(* IEC 61131-3 sources: rusty/tests/lit/single/exit, 39 files *)

(* ---- fb_exit_in_class.st ---- *)
// RUN: %COMPILE %s && %RUN | %CHECK %s
// A class can declare `FB_EXIT`. It runs for each instance when the application ends.
CLASS Logger
    METHOD FB_EXIT
        printf('logger$N');
    END_METHOD
END_CLASS

VAR_GLOBAL
    logger: Logger;
END_VAR

FUNCTION main: DINT
    printf('main done$N');
    // CHECK: main done
    // CHECK-NEXT: logger
    // CHECK-NOT: logger
END_FUNCTION

(* ---- array_elements_ascending.st ---- *)
// RUN: %COMPILE %s && %RUN | %CHECK %s
// The elements of an array are exited in ascending index order. The arrays themselves follow
// the reverse declaration order.
FUNCTION_BLOCK Slot
    VAR
        id: DINT;
    END_VAR

    METHOD FB_EXIT
        printf('slot %d$N', id);
    END_METHOD
END_FUNCTION_BLOCK

VAR_GLOBAL
    first: ARRAY[0..1] OF Slot := [(id := 1), (id := 2)];
    second: ARRAY[0..1] OF Slot := [(id := 3), (id := 4)];
END_VAR

FUNCTION main: DINT
    printf('main done$N');
    // CHECK: main done
    // CHECK-NEXT: slot 3
    // CHECK-NEXT: slot 4
    // CHECK-NEXT: slot 1
    // CHECK-NEXT: slot 2
    // CHECK-NOT: slot
END_FUNCTION

(* ---- array_with_negative_lower_bound.st ---- *)
// RUN: %COMPILE %s && %RUN | %CHECK %s
// An array whose range goes from a negative to a positive index is exited from its lowest
// index to its highest index. Each element prints its own index.
FUNCTION_BLOCK Slot
    VAR
        index: DINT;
    END_VAR

    METHOD FB_EXIT
        printf('slot %d$N', index);
    END_METHOD
END_FUNCTION_BLOCK

VAR_GLOBAL
    slots: ARRAY[-2..4] OF Slot;
END_VAR

FUNCTION main: DINT
    VAR
        i: DINT;
    END_VAR

    FOR i := -2 TO 4 DO
        slots[i].index := i;
    END_FOR

    printf('main done$N');
    // CHECK: main done
    // CHECK-NEXT: slot -2
    // CHECK-NEXT: slot -1
    // CHECK-NEXT: slot 0
    // CHECK-NEXT: slot 1
    // CHECK-NEXT: slot 2
    // CHECK-NEXT: slot 3
    // CHECK-NEXT: slot 4
    // CHECK-NOT: slot
END_FUNCTION

(* ---- array_with_two_dimensions.st ---- *)
// RUN: %COMPILE %s && %RUN | %CHECK %s
// The elements of an array with two dimensions are exited row by row: the last index changes
// first.
FUNCTION_BLOCK Slot
    VAR
        id: DINT;
    END_VAR

    METHOD FB_EXIT
        printf('slot %d$N', id);
    END_METHOD
END_FUNCTION_BLOCK

VAR_GLOBAL
    grid: ARRAY[1..2, 1..2] OF Slot;
END_VAR

FUNCTION main: DINT
    grid[1, 1].id := 11;
    grid[1, 2].id := 12;
    grid[2, 1].id := 21;
    grid[2, 2].id := 22;

    printf('main done$N');
    // CHECK: main done
    // CHECK-NEXT: slot 11
    // CHECK-NEXT: slot 12
    // CHECK-NEXT: slot 21
    // CHECK-NEXT: slot 22
    // CHECK-NOT: slot
END_FUNCTION

(* ---- container_before_members.st ---- *)
// RUN: %COMPILE %s && %RUN | %CHECK %s
// A function block runs its own `FB_EXIT` first, before any of its members is exited. The
// members follow in reverse declaration order.
FUNCTION_BLOCK Part
    VAR
        id: DINT;
    END_VAR

    METHOD FB_EXIT
        printf('part %d$N', id);
    END_METHOD
END_FUNCTION_BLOCK

FUNCTION_BLOCK Machine
    VAR
        first: Part := (id := 1);
        second: Part := (id := 2);
    END_VAR

    METHOD FB_EXIT
        printf('machine$N');
    END_METHOD
END_FUNCTION_BLOCK

VAR_GLOBAL
    machine: Machine;
END_VAR

FUNCTION main: DINT
    printf('main done$N');
    // CHECK: main done
    // CHECK-NEXT: machine
    // CHECK-NEXT: part 2
    // CHECK-NEXT: part 1
    // CHECK-NOT: {{machine|part}}
END_FUNCTION

(* ---- container_without_fb_exit.st ---- *)
// RUN: %COMPILE %s && %RUN | %CHECK %s
// A member is exited also when the function blocks that hold it declare no `FB_EXIT`, over
// more than one level.
FUNCTION_BLOCK Part
    METHOD FB_EXIT
        printf('part$N');
    END_METHOD
END_FUNCTION_BLOCK

FUNCTION_BLOCK Holder
    VAR
        part: Part;
    END_VAR
END_FUNCTION_BLOCK

FUNCTION_BLOCK Outer
    VAR
        holder: Holder;
    END_VAR
END_FUNCTION_BLOCK

VAR_GLOBAL
    outer: Outer;
END_VAR

FUNCTION main: DINT
    printf('main done$N');
    // CHECK: main done
    // CHECK-NEXT: part
    // CHECK-NOT: part
END_FUNCTION

(* ---- copy_by_assignment.st ---- *)
// RUN: %COMPILE %s && %RUN | %CHECK %s
// An assignment copies an instance with no call of `FB_INIT` or `FB_EXIT`. Each variable is
// exited one time, with the data it holds at that moment.
FUNCTION_BLOCK Token
    VAR
        id: DINT;
    END_VAR

    METHOD FB_EXIT
        printf('exit %d$N', id);
    END_METHOD
END_FUNCTION_BLOCK

VAR_GLOBAL
    target: Token := (id := 1);
    source: Token := (id := 2);
END_VAR

FUNCTION main: DINT
    target := source;
    printf('assigned$N');
    printf('main done$N');
    // CHECK: assigned
    // CHECK-NEXT: main done
    // CHECK-NEXT: exit 2
    // CHECK-NEXT: exit 2
    // CHECK-NOT: exit
END_FUNCTION

(* ---- copy_by_value_input.st ---- *)
// RUN: %COMPILE %s && %RUN | %CHECK %s
// An input that is passed by value is a copy of the argument, made with no call of `FB_INIT`.
// The copy is not exited at the end of the call. The argument is exited one time, when the
// application ends.
FUNCTION_BLOCK Token
    VAR
        id: DINT;
    END_VAR

    METHOD FB_EXIT
        printf('exit %d$N', id);
    END_METHOD
END_FUNCTION_BLOCK

FUNCTION inspect: DINT
    VAR_INPUT
        copy: Token;
    END_VAR

    printf('inspect %d$N', copy.id);
END_FUNCTION

VAR_GLOBAL
    source: Token := (id := 1);
END_VAR

FUNCTION main: DINT
    inspect(source);
    printf('main done$N');
    // CHECK: inspect 1
    // CHECK-NEXT: main done
    // CHECK-NEXT: exit 1
    // CHECK-NOT: exit
END_FUNCTION

(* ---- early_return_case.st ---- *)
// RUN: %COMPILE %s && %RUN | %CHECK %s
// A local instance is exited when the call leaves the body through a `RETURN` in a `CASE` branch.
// The statements after the `RETURN` do not run.
FUNCTION_BLOCK Guard
    METHOD FB_EXIT
        printf('exit$N');
    END_METHOD
END_FUNCTION_BLOCK

FUNCTION work: DINT
    VAR
        guard: Guard;
    END_VAR

    CASE 1 OF
        1: RETURN;
    END_CASE
    printf('not reached$N');
END_FUNCTION

FUNCTION main: DINT
    work();
    printf('main done$N');
    // CHECK-NOT: not reached
    // CHECK: exit
    // CHECK-NEXT: main done
    // CHECK-NOT: exit
END_FUNCTION

(* ---- early_return_for.st ---- *)
// RUN: %COMPILE %s && %RUN | %CHECK %s
// A local instance is exited when the call leaves the body through a `RETURN` in a `FOR` loop.
// The statements after the `RETURN` do not run.
FUNCTION_BLOCK Guard
    METHOD FB_EXIT
        printf('exit$N');
    END_METHOD
END_FUNCTION_BLOCK

FUNCTION work: DINT
    VAR
        guard: Guard;
        i: DINT;
    END_VAR

    FOR i := 0 TO 5 DO
        RETURN;
    END_FOR
    printf('not reached$N');
END_FUNCTION

FUNCTION main: DINT
    work();
    printf('main done$N');
    // CHECK-NOT: not reached
    // CHECK: exit
    // CHECK-NEXT: main done
    // CHECK-NOT: exit
END_FUNCTION

(* ---- early_return_if.st ---- *)
// RUN: %COMPILE %s && %RUN | %CHECK %s
// A local instance is exited when the call leaves the body through a `RETURN` in an `IF` branch.
// The statements after the `RETURN` do not run.
FUNCTION_BLOCK Guard
    METHOD FB_EXIT
        printf('exit$N');
    END_METHOD
END_FUNCTION_BLOCK

FUNCTION work: DINT
    VAR
        guard: Guard;
    END_VAR

    IF TRUE THEN
        RETURN;
    END_IF
    printf('not reached$N');
END_FUNCTION

FUNCTION main: DINT
    work();
    printf('main done$N');
    // CHECK-NOT: not reached
    // CHECK: exit
    // CHECK-NEXT: main done
    // CHECK-NOT: exit
END_FUNCTION

(* ---- early_return_repeat.st ---- *)
// RUN: %COMPILE %s && %RUN | %CHECK %s
// A local instance is exited when the call leaves the body through a `RETURN` in a `REPEAT` loop.
// The statements after the `RETURN` do not run.
FUNCTION_BLOCK Guard
    METHOD FB_EXIT
        printf('exit$N');
    END_METHOD
END_FUNCTION_BLOCK

FUNCTION work: DINT
    VAR
        guard: Guard;
    END_VAR

    REPEAT
        RETURN;
    UNTIL TRUE END_REPEAT
    printf('not reached$N');
END_FUNCTION

FUNCTION main: DINT
    work();
    printf('main done$N');
    // CHECK-NOT: not reached
    // CHECK: exit
    // CHECK-NEXT: main done
    // CHECK-NOT: exit
END_FUNCTION

(* ---- early_return_top_level.st ---- *)
// RUN: %COMPILE %s && %RUN | %CHECK %s
// A local instance is exited when the call leaves the body through a `RETURN` at the top level
// of the body. The statements after the `RETURN` do not run.
FUNCTION_BLOCK Guard
    METHOD FB_EXIT
        printf('exit$N');
    END_METHOD
END_FUNCTION_BLOCK

FUNCTION work: DINT
    VAR
        guard: Guard;
    END_VAR

    RETURN;
    printf('not reached$N');
END_FUNCTION

FUNCTION main: DINT
    work();
    printf('main done$N');
    // CHECK-NOT: not reached
    // CHECK: exit
    // CHECK-NEXT: main done
    // CHECK-NOT: exit
END_FUNCTION

(* ---- early_return_while.st ---- *)
// RUN: %COMPILE %s && %RUN | %CHECK %s
// A local instance is exited when the call leaves the body through a `RETURN` in a `WHILE` loop.
// The statements after the `RETURN` do not run.
FUNCTION_BLOCK Guard
    METHOD FB_EXIT
        printf('exit$N');
    END_METHOD
END_FUNCTION_BLOCK

FUNCTION work: DINT
    VAR
        guard: Guard;
    END_VAR

    WHILE TRUE DO
        RETURN;
    END_WHILE
    printf('not reached$N');
END_FUNCTION

FUNCTION main: DINT
    work();
    printf('main done$N');
    // CHECK-NOT: not reached
    // CHECK: exit
    // CHECK-NEXT: main done
    // CHECK-NOT: exit
END_FUNCTION

(* ---- explicit_call.st ---- *)
// RUN: %COMPILE %s && %RUN | %CHECK %s
// `FB_EXIT` is a normal method for user code. A call from user code runs it, and the call at
// the end of the application follows as usual.
FUNCTION_BLOCK Token
    VAR
        id: DINT;
    END_VAR

    METHOD FB_EXIT
        printf('exit %d$N', id);
    END_METHOD
END_FUNCTION_BLOCK

VAR_GLOBAL
    token: Token := (id := 1);
END_VAR

FUNCTION main: DINT
    token.FB_EXIT();
    printf('main done$N');
    // CHECK: exit 1
    // CHECK-NEXT: main done
    // CHECK-NEXT: exit 1
    // CHECK-NOT: exit
END_FUNCTION

(* ---- fb_exit_in_program.st ---- *)
// RUN: %COMPILE %s && %RUN | %CHECK %s
// A program can declare `FB_EXIT`. It runs when the application ends, before the members of the
// program are exited.
FUNCTION_BLOCK Part
    METHOD FB_EXIT
        printf('part$N');
    END_METHOD
END_FUNCTION_BLOCK

PROGRAM prog
    VAR
        part: Part;
    END_VAR

    METHOD FB_EXIT
        printf('prog$N');
    END_METHOD
END_PROGRAM

FUNCTION main: DINT
    printf('main done$N');
    // CHECK: main done
    // CHECK-NEXT: prog
    // CHECK-NEXT: part
    // CHECK-NOT: {{prog|part}}
END_FUNCTION

(* ---- function_locals.st ---- *)
// RUN: %COMPILE %s && %RUN | %CHECK %s
// A function block instance that is local to a function is initialized at the start of each
// call and exited at the end of each call, in reverse declaration order.
FUNCTION_BLOCK Guard
    VAR
        id: DINT;
    END_VAR

    METHOD FB_EXIT
        printf('exit %d$N', id);
    END_METHOD
END_FUNCTION_BLOCK

FUNCTION work: DINT
    VAR
        first: Guard := (id := 1);
        second: Guard := (id := 2);
    END_VAR

    printf('work$N');
END_FUNCTION

FUNCTION main: DINT
    work();
    work();
    printf('main done$N');
    // CHECK: work
    // CHECK-NEXT: exit 2
    // CHECK-NEXT: exit 1
    // CHECK-NEXT: work
    // CHECK-NEXT: exit 2
    // CHECK-NEXT: exit 1
    // CHECK-NEXT: main done
    // CHECK-NOT: exit
END_FUNCTION

(* ---- function_return_value.st ---- *)
// RUN: %COMPILE %s && %RUN | %CHECK %s
// The instance that a function returns is initialized and exited on each call. The caller
// receives a copy, which is exited again with the variable that holds it.
FUNCTION_BLOCK Token
    VAR
        id: DINT;
    END_VAR

    METHOD FB_INIT
        printf('init$N');
    END_METHOD

    METHOD FB_EXIT
        printf('exit %d$N', id);
    END_METHOD
END_FUNCTION_BLOCK

FUNCTION makeToken: Token
    makeToken.id := 7;
    printf('make$N');
END_FUNCTION

VAR_GLOBAL
    kept: Token;
END_VAR

FUNCTION main: DINT
    printf('main$N');
    kept := makeToken();
    printf('main done$N');
    // CHECK: init
    // CHECK-NEXT: main
    // CHECK-NEXT: init
    // CHECK-NEXT: make
    // CHECK-NEXT: exit 7
    // CHECK-NEXT: main done
    // CHECK-NEXT: exit 7
    // CHECK-NOT: exit
END_FUNCTION

(* ---- global_and_program_instances.st ---- *)
// RUN: %COMPILE %s && %RUN | %CHECK %s
// `FB_EXIT` runs one time for each instance when the application ends. Program members are
// exited before globals, the reverse of their initialization.
FUNCTION_BLOCK Connection
    VAR
        id: DINT;
    END_VAR

    METHOD FB_INIT
        printf('init$N');
    END_METHOD

    METHOD FB_EXIT
        printf('exit %d$N', id);
    END_METHOD
END_FUNCTION_BLOCK

VAR_GLOBAL
    global: Connection := (id := 1);
END_VAR

PROGRAM prog
    VAR
        member: Connection := (id := 2);
    END_VAR
END_PROGRAM

FUNCTION main: DINT
    printf('main done$N');
    // CHECK: init
    // CHECK-NEXT: init
    // CHECK-NEXT: main done
    // CHECK-NEXT: exit 2
    // CHECK-NEXT: exit 1
    // CHECK-NOT: exit
END_FUNCTION

(* ---- inheritance_derived_before_base.st ---- *)
// RUN: %COMPILE %s && %RUN | %CHECK %s
// With inheritance, the derived level runs its `FB_EXIT` and exits its members, then the base
// level does the same. The base `FB_EXIT` runs with no explicit call.
FUNCTION_BLOCK Part
    VAR
        id: DINT;
    END_VAR

    METHOD FB_EXIT
        printf('part %d$N', id);
    END_METHOD
END_FUNCTION_BLOCK

FUNCTION_BLOCK Base
    VAR
        basePart: Part := (id := 1);
    END_VAR

    METHOD FB_EXIT
        printf('base$N');
    END_METHOD
END_FUNCTION_BLOCK

FUNCTION_BLOCK Derived EXTENDS Base
    VAR
        derivedPart: Part := (id := 2);
    END_VAR

    METHOD FB_EXIT
        printf('derived$N');
    END_METHOD
END_FUNCTION_BLOCK

VAR_GLOBAL
    instance: Derived;
END_VAR

FUNCTION main: DINT
    printf('main done$N');
    // CHECK: main done
    // CHECK-NEXT: derived
    // CHECK-NEXT: part 2
    // CHECK-NEXT: base
    // CHECK-NEXT: part 1
    // CHECK-NOT: {{derived|base|part}}
END_FUNCTION

(* ---- inheritance_fb_exit_is_inherited.st ---- *)
// RUN: %COMPILE %s && %RUN | %CHECK %s
// A function block that declares no `FB_EXIT` runs the one of its base, one time for each
// instance.
FUNCTION_BLOCK Base
    METHOD FB_EXIT
        printf('base$N');
    END_METHOD
END_FUNCTION_BLOCK

FUNCTION_BLOCK Middle EXTENDS Base
END_FUNCTION_BLOCK

VAR_GLOBAL
    middle: Middle;
END_VAR

FUNCTION main: DINT
    printf('main done$N');
    // CHECK: main done
    // CHECK-NEXT: base
    // CHECK-NOT: base
END_FUNCTION

(* ---- inheritance_level_without_fb_exit.st ---- *)
// RUN: %COMPILE %s && %RUN | %CHECK %s
// A level without `FB_EXIT` between two levels that declare it is skipped: the derived
// `FB_EXIT` runs, then the one of the base.
FUNCTION_BLOCK Base
    METHOD FB_EXIT
        printf('base$N');
    END_METHOD
END_FUNCTION_BLOCK

FUNCTION_BLOCK Middle EXTENDS Base
END_FUNCTION_BLOCK

FUNCTION_BLOCK Derived EXTENDS Middle
    METHOD FB_EXIT
        printf('derived$N');
    END_METHOD
END_FUNCTION_BLOCK

VAR_GLOBAL
    derived: Derived;
END_VAR

FUNCTION main: DINT
    printf('main done$N');
    // CHECK: main done
    // CHECK-NEXT: derived
    // CHECK-NEXT: base
    // CHECK-NOT: {{derived|base}}
END_FUNCTION

(* ---- local_array.st ---- *)
// RUN: %COMPILE %s && %RUN | %CHECK %s
// A local array of function block instances is exited at the end of the call, the elements in
// ascending order.
FUNCTION_BLOCK Guard
    VAR
        id: DINT;
    END_VAR

    METHOD FB_EXIT
        printf('exit %d$N', id);
    END_METHOD
END_FUNCTION_BLOCK

FUNCTION work: DINT
    VAR
        guards: ARRAY[0..1] OF Guard := [(id := 1), (id := 2)];
    END_VAR

    printf('work$N');
END_FUNCTION

FUNCTION main: DINT
    work();
    printf('main done$N');
    // CHECK: work
    // CHECK-NEXT: exit 1
    // CHECK-NEXT: exit 2
    // CHECK-NEXT: main done
    // CHECK-NOT: exit
END_FUNCTION

(* ---- local_struct.st ---- *)
// RUN: %COMPILE %s && %RUN | %CHECK %s
// A local struct with function block fields is exited at the end of the call, the fields in
// reverse declaration order.
FUNCTION_BLOCK Guard
    VAR
        id: DINT;
    END_VAR

    METHOD FB_EXIT
        printf('exit %d$N', id);
    END_METHOD
END_FUNCTION_BLOCK

TYPE Pair: STRUCT
    first: Guard := (id := 1);
    second: Guard := (id := 2);
END_STRUCT END_TYPE

FUNCTION work: DINT
    VAR
        pair: Pair;
    END_VAR

    printf('work$N');
END_FUNCTION

FUNCTION main: DINT
    work();
    printf('main done$N');
    // CHECK: work
    // CHECK-NEXT: exit 2
    // CHECK-NEXT: exit 1
    // CHECK-NEXT: main done
    // CHECK-NOT: exit
END_FUNCTION

(* ---- method_locals.st ---- *)
// RUN: %COMPILE %s && %RUN | %CHECK %s
// A function block instance that is local to a method is exited at the end of each call of the
// method.
FUNCTION_BLOCK Guard
    METHOD FB_EXIT
        printf('exit$N');
    END_METHOD
END_FUNCTION_BLOCK

FUNCTION_BLOCK Worker
    METHOD run
        VAR
            local: Guard;
        END_VAR

        printf('run$N');
    END_METHOD
END_FUNCTION_BLOCK

VAR_GLOBAL
    worker: Worker;
END_VAR

FUNCTION main: DINT
    worker.run();
    worker.run();
    printf('main done$N');
    // CHECK: run
    // CHECK-NEXT: exit
    // CHECK-NEXT: run
    // CHECK-NEXT: exit
    // CHECK-NEXT: main done
    // CHECK-NOT: exit
END_FUNCTION

(* ---- nested_instances_depth_first.st ---- *)
// RUN: %COMPILE %s && %RUN | %CHECK %s
// Nested instances are exited depth first: a member is exited together with the members below
// it, before the next member, and a whole instance before the next independent instance.
FUNCTION_BLOCK Leaf
    METHOD FB_EXIT
        printf('leaf$N');
    END_METHOD
END_FUNCTION_BLOCK

FUNCTION_BLOCK Branch
    VAR
        id: DINT;
        leaf: Leaf;
    END_VAR

    METHOD FB_EXIT
        printf('branch %d$N', id);
    END_METHOD
END_FUNCTION_BLOCK

FUNCTION_BLOCK Tree
    VAR
        id: DINT;
        left: Branch := (id := 1);
        right: Branch := (id := 2);
    END_VAR

    METHOD FB_EXIT
        printf('tree %d$N', id);
    END_METHOD
END_FUNCTION_BLOCK

VAR_GLOBAL
    oak: Tree := (id := 1);
    pine: Tree := (id := 2);
END_VAR

FUNCTION main: DINT
    printf('main done$N');
    // CHECK: main done
    // CHECK-NEXT: tree 2
    // CHECK-NEXT: branch 2
    // CHECK-NEXT: leaf
    // CHECK-NEXT: branch 1
    // CHECK-NEXT: leaf
    // CHECK-NEXT: tree 1
    // CHECK-NEXT: branch 2
    // CHECK-NEXT: leaf
    // CHECK-NEXT: branch 1
    // CHECK-NEXT: leaf
    // CHECK-NOT: {{tree|branch|leaf}}
END_FUNCTION

(* ---- not_owned_pointer.st ---- *)
// RUN: %COMPILE %s && %RUN | %CHECK %s
// A pointer refers to an instance that is owned elsewhere. It causes no additional `FB_EXIT`:
// the one instance is exited one time.
FUNCTION_BLOCK Slot
    METHOD FB_EXIT
        printf('slot$N');
    END_METHOD
END_FUNCTION_BLOCK

FUNCTION_BLOCK User
    VAR
        ptr: REF_TO Slot := REF(shared);
    END_VAR
END_FUNCTION_BLOCK

VAR_GLOBAL
    shared: Slot;
    ptr: REF_TO Slot := REF(shared);
    user: User;
END_VAR

FUNCTION main: DINT
    printf('main done$N');
    // CHECK: main done
    // CHECK-NEXT: slot
    // CHECK-NOT: slot
END_FUNCTION

(* ---- not_owned_reference.st ---- *)
// RUN: %COMPILE %s && %RUN | %CHECK %s
// A reference refers to an instance that is owned elsewhere. It causes no additional `FB_EXIT`:
// the one instance is exited one time.
FUNCTION_BLOCK Slot
    METHOD FB_EXIT
        printf('slot$N');
    END_METHOD
END_FUNCTION_BLOCK

FUNCTION_BLOCK User
    VAR
        reference: REFERENCE TO Slot REF= shared;
    END_VAR
END_FUNCTION_BLOCK

VAR_GLOBAL
    shared: Slot;
    reference: REFERENCE TO Slot REF= shared;
    user: User;
END_VAR

FUNCTION main: DINT
    printf('main done$N');
    // CHECK: main done
    // CHECK-NEXT: slot
    // CHECK-NOT: slot
END_FUNCTION

(* ---- not_owned_var_in_out.st ---- *)
// RUN: %COMPILE %s && %RUN | %CHECK %s
// A `VAR_IN_OUT` of a function block or a function refers to an instance of the caller. It
// causes no additional `FB_EXIT`: the one instance is exited one time.
FUNCTION_BLOCK Slot
    METHOD FB_EXIT
        printf('slot$N');
    END_METHOD
END_FUNCTION_BLOCK

FUNCTION_BLOCK User
    VAR_IN_OUT
        borrowed: Slot;
    END_VAR
END_FUNCTION_BLOCK

FUNCTION borrow: DINT
    VAR_IN_OUT
        borrowed: Slot;
    END_VAR
END_FUNCTION

VAR_GLOBAL
    shared: Slot;
    user: User;
END_VAR

FUNCTION main: DINT
    user(borrowed := shared);
    borrow(shared);
    printf('main done$N');
    // CHECK: main done
    // CHECK-NEXT: slot
    // CHECK-NOT: slot
END_FUNCTION

(* ---- recursion.st ---- *)
// RUN: %COMPILE %s && %RUN | %CHECK %s
// Each level of a recursion has its own local instance, which is exited when that level returns.
FUNCTION_BLOCK Guard
    VAR
        id: DINT;
    END_VAR

    METHOD FB_EXIT
        printf('exit %d$N', id);
    END_METHOD
END_FUNCTION_BLOCK

FUNCTION descend: DINT
    VAR_INPUT
        depth: DINT;
    END_VAR
    VAR
        guard: Guard;
    END_VAR

    guard.id := depth;
    IF depth < 3 THEN
        descend(depth + 1);
    END_IF
END_FUNCTION

FUNCTION main: DINT
    descend(1);
    printf('main done$N');
    // CHECK: exit 3
    // CHECK-NEXT: exit 2
    // CHECK-NEXT: exit 1
    // CHECK-NEXT: main done
    // CHECK-NOT: exit
END_FUNCTION

(* ---- reverse_declaration_order.st ---- *)
// RUN: %COMPILE %s && %RUN | %CHECK %s
// Independent instances are exited in the reverse order of their declaration, also when their
// types differ.
FUNCTION_BLOCK Motor
    VAR
        id: DINT;
    END_VAR

    METHOD FB_EXIT
        printf('motor %d$N', id);
    END_METHOD
END_FUNCTION_BLOCK

FUNCTION_BLOCK Valve
    VAR
        id: DINT;
    END_VAR

    METHOD FB_EXIT
        printf('valve %d$N', id);
    END_METHOD
END_FUNCTION_BLOCK

VAR_GLOBAL
    first: Motor := (id := 1);
    second: Valve := (id := 2);
    third: Motor := (id := 3);
END_VAR

FUNCTION main: DINT
    printf('main done$N');
    // CHECK: main done
    // CHECK-NEXT: motor 3
    // CHECK-NEXT: valve 2
    // CHECK-NEXT: motor 1
    // CHECK-NOT: {{motor|valve}}
END_FUNCTION

(* ---- signature_with_copy_code_parameter.st ---- *)
// RUN: %COMPILE %s && %RUN | %CHECK %s
// `FB_EXIT` with the input `bInCopyCode` and a `BOOL` result is called with `FALSE`.
FUNCTION_BLOCK Token
    METHOD FB_EXIT: BOOL
        VAR_INPUT
            bInCopyCode: BOOL;
        END_VAR

        IF NOT bInCopyCode THEN
            printf('exit without copy code$N');
        END_IF
    END_METHOD
END_FUNCTION_BLOCK

VAR_GLOBAL
    token: Token;
END_VAR

FUNCTION main: DINT
    printf('main done$N');
    // CHECK: main done
    // CHECK-NEXT: exit without copy code
    // CHECK-NOT: exit
END_FUNCTION

(* ---- signature_with_default_parameter.st ---- *)
// RUN: %COMPILE %s && %RUN | %CHECK %s
// `FB_EXIT` with a different signature is called with the default values of its parameters.
FUNCTION_BLOCK Counter
    METHOD FB_EXIT: DINT
        VAR_INPUT
            amount: DINT := 7;
        END_VAR

        printf('exit with amount %d$N', amount);
    END_METHOD
END_FUNCTION_BLOCK

VAR_GLOBAL
    counter: Counter;
END_VAR

FUNCTION main: DINT
    printf('main done$N');
    // CHECK: main done
    // CHECK-NEXT: exit with amount 7
    // CHECK-NOT: exit
END_FUNCTION

(* ---- struct_fields.st ---- *)
// RUN: %COMPILE %s && %RUN | %CHECK %s
// The function block fields of a struct are exited in reverse declaration order. The struct
// itself has no `FB_EXIT`, and its other fields are left alone.
FUNCTION_BLOCK Slot
    VAR
        id: DINT;
    END_VAR

    METHOD FB_EXIT
        printf('slot %d$N', id);
    END_METHOD
END_FUNCTION_BLOCK

TYPE Pair: STRUCT
    first: Slot := (id := 1);
    count: DINT;
    second: Slot := (id := 2);
END_STRUCT END_TYPE

VAR_GLOBAL
    pair: Pair;
END_VAR

FUNCTION main: DINT
    printf('main done$N');
    // CHECK: main done
    // CHECK-NEXT: slot 2
    // CHECK-NEXT: slot 1
    // CHECK-NOT: slot
END_FUNCTION

(* ---- struct_in_array.st ---- *)
// RUN: %COMPILE %s && %RUN | %CHECK %s
// A struct with a function block field is exited also when it is an array element: one time for
// each element.
FUNCTION_BLOCK Slot
    METHOD FB_EXIT
        printf('slot$N');
    END_METHOD
END_FUNCTION_BLOCK

TYPE Holder: STRUCT
    slot: Slot;
END_STRUCT END_TYPE

VAR_GLOBAL
    holders: ARRAY[0..1] OF Holder;
END_VAR

FUNCTION main: DINT
    printf('main done$N');
    // CHECK: main done
    // CHECK-NEXT: slot
    // CHECK-NEXT: slot
    // CHECK-NOT: slot
END_FUNCTION

(* ---- struct_in_function_block.st ---- *)
// RUN: %COMPILE %s && %RUN | %CHECK %s
// A struct with a function block field is exited also when it is a member of a function block.
FUNCTION_BLOCK Slot
    METHOD FB_EXIT
        printf('slot$N');
    END_METHOD
END_FUNCTION_BLOCK

TYPE Holder: STRUCT
    slot: Slot;
END_STRUCT END_TYPE

FUNCTION_BLOCK Owner
    VAR
        holder: Holder;
    END_VAR
END_FUNCTION_BLOCK

VAR_GLOBAL
    owner: Owner;
END_VAR

FUNCTION main: DINT
    printf('main done$N');
    // CHECK: main done
    // CHECK-NEXT: slot
    // CHECK-NOT: slot
END_FUNCTION

(* ---- struct_in_struct.st ---- *)
// RUN: %COMPILE %s && %RUN | %CHECK %s
// A struct with a function block field is exited also when it is a field of another struct.
FUNCTION_BLOCK Slot
    METHOD FB_EXIT
        printf('slot$N');
    END_METHOD
END_FUNCTION_BLOCK

TYPE Holder: STRUCT
    slot: Slot;
END_STRUCT END_TYPE

TYPE Wrapper: STRUCT
    holder: Holder;
END_STRUCT END_TYPE

VAR_GLOBAL
    wrapper: Wrapper;
END_VAR

FUNCTION main: DINT
    printf('main done$N');
    // CHECK: main done
    // CHECK-NEXT: slot
    // CHECK-NOT: slot
END_FUNCTION

(* ---- temporary_in_function_block.st ---- *)
// RUN: %COMPILE %s && %RUN | %CHECK %s
// A `VAR_TEMP` instance of a function block is exited at the end of each call. A member in `VAR`
// lives as long as its instance and is exited when the application ends.
FUNCTION_BLOCK Guard
    VAR
        id: DINT;
    END_VAR

    METHOD FB_EXIT
        printf('exit %d$N', id);
    END_METHOD
END_FUNCTION_BLOCK

FUNCTION_BLOCK Worker
    VAR
        member: Guard := (id := 1);
    END_VAR
    VAR_TEMP
        temporary: Guard := (id := 2);
    END_VAR

    printf('worker$N');
END_FUNCTION_BLOCK

VAR_GLOBAL
    worker: Worker;
END_VAR

FUNCTION main: DINT
    worker();
    printf('main done$N');
    // CHECK: worker
    // CHECK-NEXT: exit 2
    // CHECK-NEXT: main done
    // CHECK-NEXT: exit 1
    // CHECK-NOT: exit
END_FUNCTION

(* ---- temporary_in_program.st ---- *)
// RUN: %COMPILE %s && %RUN | %CHECK %s
// A `VAR_TEMP` instance of a program is exited at the end of each call.
FUNCTION_BLOCK Guard
    METHOD FB_EXIT
        printf('exit$N');
    END_METHOD
END_FUNCTION_BLOCK

PROGRAM prog
    VAR_TEMP
        temporary: Guard;
    END_VAR

    printf('prog$N');
END_PROGRAM

FUNCTION main: DINT
    prog();
    printf('main done$N');
    // CHECK: prog
    // CHECK-NEXT: exit
    // CHECK-NEXT: main done
    // CHECK-NOT: exit
END_FUNCTION
